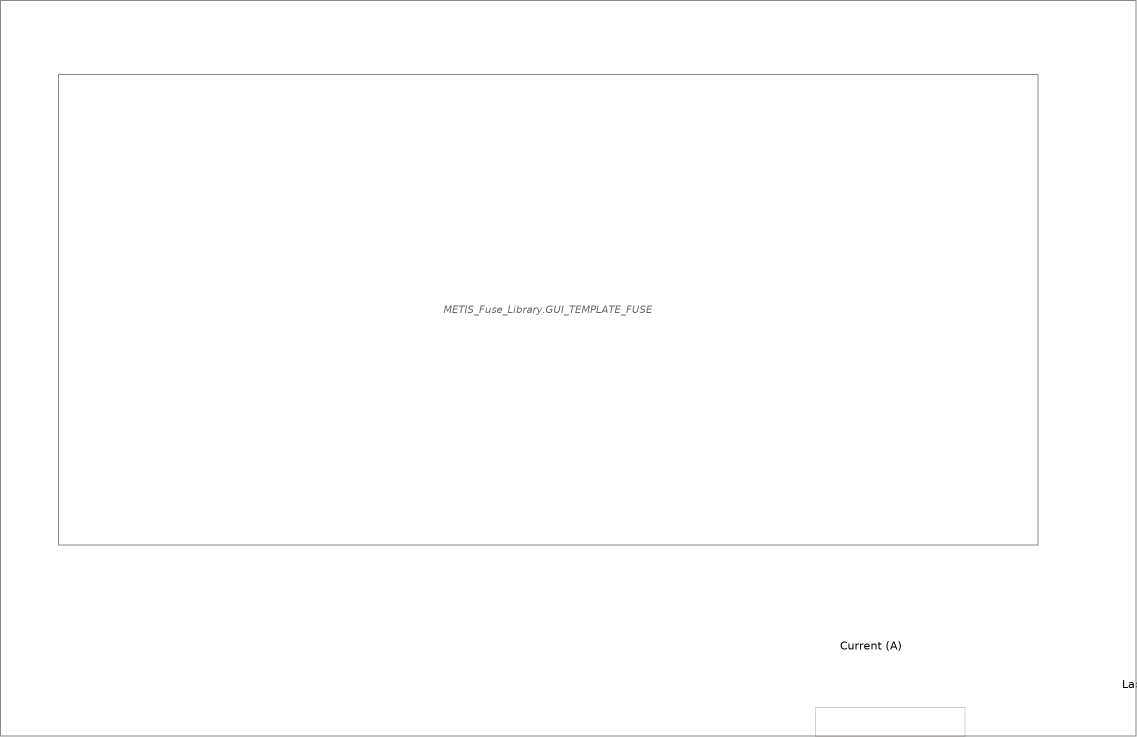
VISUALIZATION VISU_DETECTOR_POWER  // 1137x737
    Frame (58,74 980x471)
        shows METIS_Fuse_Library.GUI_TEMPLATE_FUSE(m_Instance := MAIN.nott_detector_power.fuseDetectorPower)
    Label (1137,684 0x1), "Label"
    Label (796,631 150x30), "Current (A)"
    Textfield (815,707 150x30), text variable: MAIN.nott_detector_power.lrActCurrent
END_VISUALIZATION

(* stored: Version 1.1.0.1, ProductVersion 3.1.4026.20
   Visu VISU_DETECTOR_POWER: Id {fd78a343-3473-480b-a3e2-bce600d4bcbd} *)
